(* IEC 61131-3 sources: veristc/veri-stc/tests/st-examples/feature-probes, 13 files *)

(* ---- p13_in_out_alias.st ---- *)
(* p13: VAR_IN_OUT 逐引用别名——端口是调用方存储的别名，不是副本
   场景: shared 为全局累加器；i1/i2 两个实例的 ACC 端口都绑定 shared，
         体内 LAST := ACC（读别名）+ ACC := ACC + K（写别名）。
         每周期 i1 加 tick、i2 加 100 ⇒ shared 单点跨实例累加；
         两实例 LAST 互不相同 ⇒ 实例数据仍分离。 *)
VAR_GLOBAL
  shared : DINT;
  i1 : ACCUM;
  i2 : ACCUM;
END_VAR

FUNCTION_BLOCK ACCUM
VAR_INPUT
  K : DINT;
END_VAR
VAR_OUTPUT
  LAST : DINT;
END_VAR
VAR_IN_OUT
  ACC : DINT;
END_VAR
  LAST := ACC;
  ACC := ACC + K;
END_FUNCTION_BLOCK

PROGRAM MAIN
VAR
  tick : DINT;
END_VAR
  tick := CycleCounter();
  i1(ACC := shared, K := tick);
  i2(ACC := shared, K := 100);
  PRINT('p13 shared=', shared, ' i1=', i1.LAST, ' i2=', i2.LAST, '\n');
END_PROGRAM

(* ---- p01_case.st ---- *)
(* p01: CASE 语句——单值/多值/范围/ELSE 四类分支（desugar → IF 链） *)
PROGRAM MAIN
VAR
  tick : DINT;
  code : DINT;
END_VAR
  tick := CycleCounter();
  code := 0;
  CASE tick OF
    1:
      code := 10;
    2,3:
      code := 20;
    4..6:
      code := 30;
  ELSE:
    code := 99;
  END_CASE;
  PRINT('p01 code=', code, '\n');
END_PROGRAM

(* ---- p02_for.st ---- *)
(* p02: FOR 循环——常量上界/步长/嵌套（desugar → WHILE 计数模式） *)
PROGRAM MAIN
VAR
  i : INT;      (* 类型检查规则 TS_for_int: 循环变量必须为 INT *)
  j : INT;
  sum : DINT;
  step_sum : DINT;
  pairs : DINT;
END_VAR
  sum := 0;
  FOR i := 1 TO 5 DO
    sum := sum + i;
  END_FOR;

  step_sum := 0;
  FOR i := 2 TO 8 BY 2 DO
    step_sum := step_sum + i;
  END_FOR;

  pairs := 0;
  FOR i := 1 TO 3 DO
    FOR j := 1 TO 4 DO
      pairs := pairs + 1;
    END_FOR;
  END_FOR;

  PRINT('p02 s=', sum, ' ss=', step_sum, ' c=', pairs, '\n');
END_PROGRAM

(* ---- p03_while_repeat.st ---- *)
(* p03: WHILE 递减收敛 + REPEAT-UNTIL 至少执行一次语义 *)
PROGRAM MAIN
VAR
  n : DINT;
  k : DINT;
  m : DINT;
END_VAR
  n := 100;
  k := 0;
  WHILE n > 50 DO
    n := n - 7;
    k := k + 1;
  END_WHILE;

  m := 0;
  REPEAT
    m := m + 3;
  UNTIL m >= 20
  END_REPEAT;

  PRINT('p03 n=', n, ' k=', k, ' m=', m, '\n');
END_PROGRAM

(* ---- p04_div_mod.st ---- *)
(* p04: 有符号除法/取余——负操作数截断语义（对齐 C 与 Coq Z.div/Z.rem） *)
PROGRAM MAIN
VAR
  tick : DINT;
  a : DINT;
  r : DINT;
  q : DINT;
  ne : DINT;
  nd : DINT;
  nr : DINT;
END_VAR
  tick := CycleCounter();
  a := tick * 7 + 3;
  r := a MOD 5;
  q := a / 5;
  ne := 0 - 17;
  nd := ne / 5;
  nr := ne MOD 5;
  PRINT('p04 a=', a, ' r=', r, ' q=', q, ' nd=', nd, ' nr=', nr, '\n');
END_PROGRAM

(* ---- p05_xor_bits.st ---- *)
(* p05: 布尔 XOR + 算术法位抽取。
   注：T_And/T_Or/T_Xor 形式规则仅接受 BOOL 操作数——WORD 位与在实编译管线
   不可用（safeasm-spec 声明支持、类型规则未放行，矛盾记录见 README）；
   工程惯用 / MOD 做位域抽取。ABS 因 LOCAL_SET 255 越界静默丢弃，另立项。 *)
PROGRAM MAIN
VAR
  tick : DINT;
  x : DINT;
  b : BOOL;     (* BOOL 域 XOR；BOOL→DINT 赋值被类型检查器拒绝 *)
  v : DINT;
  hi : DINT;
  lo : DINT;
  c : BOOL;
END_VAR
  tick := CycleCounter();
  x := tick * 3;
  b := (x > 5) XOR (12 > 8);
  v := tick * 65536 + 4096;
  hi := (v / 256) MOD 256;
  lo := v MOD 256;
  c := b AND (hi = 16);
  PRINT('p05 b=', b, ' hi=', hi, ' lo=', lo, ' c=', c, '\n');
END_PROGRAM

(* ---- p06_latch_state.st ---- *)
(* p06: 跨周期锁存状态——VAR_GLOBAL 持久 + 迟滞整定 + 手动复位
   场景: x = tick*25; 跳闸阈值 x>100; 复位脉冲 tick=7 *)
VAR_GLOBAL
  latched : BOOL;
END_VAR

PROGRAM MAIN
VAR
  tick : DINT;
  x : DINT;
  rst : BOOL;
END_VAR
  tick := CycleCounter();
  x := tick * 25;
  rst := tick = 7;

  latched := (NOT rst) AND ((x > 100) OR (latched AND NOT (x < 80)));
  PRINT('p06 x=', x, ' latched=', latched, '\n');
END_PROGRAM

(* ---- p07_real_arith.st ---- *)
(* p07 [XFAIL-后端缺口]: REAL 浮点算术。
   REAL 字面量自 v1.5.4 起可写也可落盘（lexer.v 十进制快路 + 主机侧立即数真值，
   已由 compiler-tests/positive/real_literals.st 逐条核对位模式）。
   但 spec 要求 F32_ADD/F32_CMP 类型导向降级；当前 global_codegen.v 的
   compile_expr_g（PROGRAM 体专用）对一切二元运算统一发 I32 指令 → 结果必然错误。
   期望 ok=1。 *)
PROGRAM MAIN
VAR
  a : REAL;
  b : REAL;
  ok : DINT;
END_VAR
  a := 1.5;
  b := a + 2.25;
  ok := 0;
  IF (b > 3.5) AND (b < 4.0) THEN
    ok := 1;
  END_IF;
  PRINT('p07 ok=', ok, '\n');
END_PROGRAM

(* ---- p08_lint_arith.st ---- *)
(* p08 [XFAIL-后端缺口]: LINT 64 位算术。
   spec 要求 I64_ADD/I64_DIV_S/I64_CMP；当前后端全部 I32 截断。
   判据用"除以 1e9 后是否等于 6"：I32 截断路径下 (a+b) mod 2^32 是环同态，
   大小比较两侧同余截断仍为真（弱判据）；除法不保持同余，能区分 64 位与
   截断路径（截断: 1705032704/1000000000 = 1 ≠ 6）。期望 ok=1。 *)
PROGRAM MAIN
VAR
  big : LINT;
  sum : LINT;
  scale : LINT;
  ok : DINT;
END_VAR
  big := 3000000000;
  sum := big + big;
  scale := sum / 1000000000;
  ok := 0;
  IF scale = 6 THEN
    ok := 1;
  END_IF;
  PRINT('p08 ok=', ok, '\n');
END_PROGRAM

(* ---- p09_array_ops.st ---- *)
(* p09 [XFAIL-后端缺口]: 静态数组读写。
   spec: 地址 = base + (idx-low)*width；当前 CS_ARRAY_ASSIGN/CE_ARRAY_ACCESS
   把数组变量当"值"再 +idx（无宽度缩放，全局数组读到的是内容不是地址）。
   期望 s=20。 *)
PROGRAM MAIN
VAR
  buf : ARRAY[0..3] OF DINT;
  i : DINT;
  s : DINT;
END_VAR
  FOR i := 0 TO 3 DO
    buf[i] := i * 10;
  END_FOR;
  s := buf[0] + buf[2];
  PRINT('p09 s=', s, '\n');
END_PROGRAM

(* ---- p10_quality_ops.st ---- *)
(* p10 [XFAIL-后端缺口]: 质量算子与质量传播。
   spec: Q_WITH(TRUE,BAD) 构造坏质量值，Q_GOOD 应为 FALSE。
   当前 CE_QUALITY_OP 仅透传数值参数，质量语义在实编译后端不存在 → 输出 1。
   期望 g=0。 *)
PROGRAM MAIN
VAR
  q : QBOOL;
  g : DINT;
END_VAR
  q := Q_WITH(TRUE, BAD);
  g := 0;
  IF Q_GOOD(q) THEN
    g := 1;
  END_IF;
  PRINT('p10 g=', g, '\n');
END_PROGRAM

(* ---- p11_nested_fn.st ---- *)
(* p11: FUNCTION 嵌套内联——Quad 调用 Twice，两层展开后与 4*tick 恒等 *)
FUNCTION Twice : DINT
VAR_INPUT
  x : DINT;
END_VAR
  Twice := x + x;
END_FUNCTION

FUNCTION Quad : DINT
VAR_INPUT
  x : DINT;
END_VAR
  Quad := Twice(Twice(x));
END_FUNCTION

PROGRAM MAIN
VAR
  tick : DINT;
  q : DINT;
  diff : DINT;
END_VAR
  tick := CycleCounter();
  q := Quad(tick);
  diff := q - 4 * tick;
  PRINT('p11 q=', q, ' diff=', diff, '\n');
END_PROGRAM

(* ---- p12_divzero_trap.st ---- *)
(* p12: 除零运行时陷阱——tick=3 时触发 10/0，期望 VM 报错退出，
   前两个周期正常输出 e=10 *)
PROGRAM MAIN
VAR
  tick : DINT;
  e : DINT;
END_VAR
  tick := CycleCounter();
  e := 10;
  IF tick = 3 THEN
    e := e / 0;
  END_IF;
  PRINT('p12 e=', e, '\n');
END_PROGRAM
